(* IEC 61131-3 sources: rusty/tests/lit/single/functions, 19 files *)

(* ---- output_aggregate_initializers.st ---- *)
// RUN: %COMPILE %s && %RUN | %CHECK %s
// A struct literal, an array literal, and a string on a VAR_OUTPUT are applied by the lowered
// stack initializer of the function; the entry reset only zero-fills aggregates.
TYPE S : STRUCT
    x : INT;
    y : INT;
END_STRUCT END_TYPE

FUNCTION f
    VAR_OUTPUT
        out : S := (x := 7);
        arr : ARRAY[0..1] OF INT := [1, 2];
        s : STRING := 'abc';
    END_VAR
END_FUNCTION

FUNCTION main
    VAR
        v : S;
        a : ARRAY[0..1] OF INT;
        str : STRING;
    END_VAR
    v.y := 5;
    f(out => v, arr => a, s => str);
    printf('v = (%d, %d), a = [%d, %d], s = %s$N', v.x, v.y, a[0], a[1], str);
    // CHECK: v = (7, 0), a = [1, 2], s = abc
END_FUNCTION

(* ---- by_ref_argument_is_evaluated_once.st ---- *)
// RUN: %COMPILE %s && %RUN | %CHECK %s
// An expression passed to a by-reference input is evaluated once, also when the compiler carries it
// out through a replacement such as a builtin or a standard library call

VAR_GLOBAL
    calls : DINT;
END_VAR

FUNCTION next_number : DINT
    calls := calls + 1;
    next_number := calls;
END_FUNCTION

FUNCTION next_duration : TIME
    calls := calls + 1;
    next_duration := T#5s;
END_FUNCTION

FUNCTION read_number : DINT
VAR_INPUT {ref}
    in : DINT;
END_VAR
    read_number := in;
END_FUNCTION

FUNCTION read_duration : TIME
VAR_INPUT {ref}
    in : TIME;
END_VAR
    read_duration := in;
END_FUNCTION

FUNCTION main : DINT
    VAR
        n : DINT := 10;
        t : TIME := T#1s;
        result : DINT;
        duration : TIME;
    END_VAR

    result := read_number(n + next_number());
    printf('%d$N', result);                                                         // CHECK: 11
    printf('%d$N', calls);                                                          // CHECK: 1

    result := read_number(ADD(n, next_number()));
    printf('%d$N', result);                                                         // CHECK: 12
    printf('%d$N', calls);                                                          // CHECK: 2

    duration := read_duration(ADD(t, next_duration()));
    printf('%s$N', REF(TIME_TO_STRING(duration)));                                  // CHECK: T#6s
    printf('%d$N', calls);                                                          // CHECK: 3

END_FUNCTION

(* ---- call_with_array_access_on_result.st ---- *)
// RUN: %COMPILE %s && %RUN | %CHECK %s

FUNCTION foo: ARRAY[1..5] OF DINT
    foo := [5, 4, 3, 2, 1];
END_FUNCTION

FUNCTION alwaysOne: DINT
    alwaysOne := 1;
END_FUNCTION

FUNCTION main
    VAR
        value: DINT;
        one: DINT := 1;
        two: DINT := 2;
    END_VAR

    // CHECK: 5
    value := foo()[1];
    printf('%d$N', value);

    // CHECK: 3
    value := foo()[1 + 2];
    printf('%d$N', value);

    // CHECK: 5
    value := foo()[one];
    printf('%d$N', value);

    // CHECK: 3
    value := foo()[one + two];
    printf('%d$N', value);

    // CHECK: 5
    value := foo()[alwaysOne()];
    printf('%d$N', value);
END_FUNCTION

(* ---- deeply_nested_calls.st ---- *)
// RUN: %COMPILE %s && %RUN | %CHECK %s
// Deeply nested calls compile in time linear to their depth

FUNCTION increment : DINT
    VAR_INPUT
        value : DINT;
    END_VAR

    increment := value + 1;
END_FUNCTION

FUNCTION main
    VAR
        x : DINT := 0;
    END_VAR

    x := increment(increment(increment(increment(increment(increment(increment(increment(increment(increment(increment(increment(increment(increment(increment(increment(increment(increment(increment(increment(increment(increment(increment(increment(increment(increment(increment(increment(increment(increment(x))))))))))))))))))))))))))))));
    printf('%d$N', x);                                                              // CHECK: 30

END_FUNCTION

(* ---- default_params.st ---- *)
// RUN: %COMPILE %s && %RUN | %CHECK %s
FUNCTION func : int
  VAR_INPUT
    in : INT := 42;
  END_VAR
  func := in;
END_FUNCTION

FUNCTION main : DINT

    PRINTF('func complete:%d$N', func(13)); //CHECK: func complete:13
    PRINTF('func incomplete:%d$N', func()); //CHECK: func incomplete:42

END_FUNCTION

(* ---- function_output_should_be_cast_if_needed.st ---- *)
// RUN: %COMPILE %s && %RUN | %CHECK %s
FUNCTION outputCastIntToReal : INT
    VAR_OUTPUT
        result : REAL;
    END_VAR

    result := 42.0;
END_FUNCTION

FUNCTION outputNoCastInt : INT
    VAR_OUTPUT
        result : INT;
    END_VAR

    result := 52;
END_FUNCTION

FUNCTION outputCastRealToInt : INT
    VAR_OUTPUT
        result : INT;
    END_VAR

    result := 62;
END_FUNCTION

FUNCTION outputNoCastReal : INT
    VAR_OUTPUT
        result : REAL;
    END_VAR

    result := 72.0;
END_FUNCTION

FUNCTION main
    VAR
        i1 : INT;
        i2 : INT;
        r1 : REAL;
        r2 : REAL;
    END_VAR

    i1 := 31;
    i2 := 32;
    r1 := 33;
    r2 := 34;

    // ----------------- //
    // -- INT to REAL -- //

    outputCastIntToReal(
        result => i1
    );

    // CHECK: 42
    PRINTF('%d$N', i1);

    // ---------------- //
    // -- INT to INT -- //

    outputNoCastInt(
        result => i2
    );

    // CHECK: 52
    PRINTF('%d$N', i2);

    // ----------------- //
    // -- REAL to INT -- //

    outputCastRealToInt(
        result => r1
    );

    // CHECK: 62.0
    PRINTF('%.1f$N', r1);

    // ------------------ //
    // -- REAL to REAL -- //

    outputNoCastReal(
        result => r2
    );

    // CHECK: 72.0
    PRINTF('%.1f$N', r2);
END_FUNCTION

(* ---- function_parameter_with_bit_access.st ---- *)
// RUN: %COMPILE %s && %RUN | %CHECK %s
FUNCTION FLIP
    VAR_INPUT
        in: BYTE;
    END_VAR
    VAR_OUTPUT
        out : BYTE;
    END_VAR
    out := NOT(in);
END_FUNCTION

FUNCTION main
    VAR
        wordVar : WORD;
    END_VAR

    wordVar := 0;
    FLIP(2#01010101, wordVar.%b0);

    // CHECK: wordVar=170
    PRINTF('wordVar=%d$N', wordVar);
END_FUNCTION

(* ---- function_parameter_with_bit_access_named_params.st ---- *)
// RUN: %COMPILE %s && %RUN | %CHECK %s
FUNCTION FLIP
    VAR_INPUT
        in: BYTE;
    END_VAR
    VAR_OUTPUT
        out : BYTE;
    END_VAR
    out := NOT(in);
END_FUNCTION

FUNCTION main
    VAR
        wordVar : WORD;
    END_VAR

    wordVar := 0;
    FLIP(in := 2#01010101, out => wordVar.%b0);

    // CHECK: wordVar=170
    PRINTF('wordVar=%d$N', wordVar);
END_FUNCTION

(* ---- output_reset_on_every_call.st ---- *)
// RUN: %COMPILE %s && %RUN | %CHECK %s
// A function output that a path does not assign comes back at its default on every call, not at
// the value a previous call left in the caller's variable.
FUNCTION clamp_flag
    VAR_INPUT
        value : INT;
    END_VAR
    VAR_OUTPUT
        too_big : BOOL;
    END_VAR
    IF value > 2 THEN
        too_big := TRUE;
    END_IF
END_FUNCTION

FUNCTION main
    VAR
        i : INT;
        flag : BOOL;
    END_VAR
    FOR i := 1 TO 5 DO
        clamp_flag(i, flag);
        printf('%d: %d$N', i, flag);
    END_FOR
    // CHECK: 1: 0
    // CHECK-NEXT: 2: 0
    // CHECK-NEXT: 3: 1
    // CHECK-NEXT: 4: 1
    // CHECK-NEXT: 5: 1
    flag := TRUE;
    clamp_flag(1, flag);
    printf('after: %d$N', flag);
    // CHECK-NEXT: after: 0
END_FUNCTION

(* ---- function_block_output_should_be_cast_if_needed.st ---- *)
// RUN: %COMPILE %s && %RUN | %CHECK %s
FUNCTION_BLOCK outputCastIntToReal_fb
    VAR_OUTPUT
        result : REAL;
    END_VAR

    result := 42.0;
END_FUNCTION_BLOCK

FUNCTION_BLOCK outputNoCastInt_fb
    VAR_OUTPUT
        result : INT;
    END_VAR

    result := 52;
END_FUNCTION_BLOCK

FUNCTION_BLOCK outputCastRealToInt_fb
    VAR_OUTPUT
        result : INT;
    END_VAR

    result := 62;
END_FUNCTION_BLOCK

FUNCTION_BLOCK outputNoCastReal_fb
    VAR_OUTPUT
        result : REAL;
    END_VAR

    result := 72.0;
END_FUNCTION_BLOCK

FUNCTION main
    VAR
        outputCastIntToReal : outputCastIntToReal_fb;
        outputNoCastInt : outputNoCastInt_fb;
        outputCastRealToInt : outputCastRealToInt_fb;
        outputNoCastReal : outputNoCastReal_fb;

        i1 : INT;
        i2 : INT;
        r1 : REAL;
        r2 : REAL;
    END_VAR

    i1 := 31;
    i2 := 32;
    r1 := 33;
    r2 := 34;

    // ----------------- //
    // -- INT to REAL -- //

    outputCastIntToReal(
        result => i1
    );

    // CHECK: 42
    PRINTF('%d$N', i1);

    // ---------------- //
    // -- INT to INT -- //

    outputNoCastInt(
        result => i2
    );

    // CHECK: 52
    PRINTF('%d$N', i2);

    // ----------------- //
    // -- REAL to INT -- //

    outputCastRealToInt(
        result => r1
    );

    // CHECK: 62.0
    PRINTF('%.1f$N', r1);

    // ------------------ //
    // -- REAL to REAL -- //

    outputNoCastReal(
        result => r2
    );

    // CHECK: 72.0
    PRINTF('%.1f$N', r2);
END_FUNCTION

(* ---- function_output_to_bit_direct_access.st ---- *)
// RUN: %COMPILE %s && %RUN | %CHECK %s

// Regression test for https://github.com/PLC-lang/rusty/issues/1239
// `fun(out => bar.4)` and `myFb(out => bar.4)` previously generated IR that
// computed the bit address but never stored the function's output back into
// the underlying integer.
FUNCTION fun
    VAR_OUTPUT
        foo : BOOL;
    END_VAR
    foo := TRUE;
END_FUNCTION

FUNCTION_BLOCK fb
    VAR_OUTPUT
        foo : BOOL;
    END_VAR
    foo := TRUE;
END_FUNCTION_BLOCK

FUNCTION main : DINT
    VAR
        bar  : DINT;
        myFb : fb;
    END_VAR

    bar := 0;
    fun(foo => bar.4);
    PRINTF('after_fun=%d$N', bar);
    // CHECK: after_fun=16

    bar := 0;
    myFb(foo => bar.4);
    PRINTF('after_fb=%d$N', bar);
    // CHECK: after_fb=16

    // Non-zero seed: anchors that bits 0–3 are *preserved* when the FB output
    // writes bit 4. A regression that clobbered the integer (e.g. wrote a full
    // word instead of just the bit) would surface here as 16 instead of 17.
    bar := 1;
    myFb(foo => bar.4);
    PRINTF('after_fb_seeded=%d$N', bar);
    // CHECK: after_fb_seeded=17
END_FUNCTION

(* ---- output_pointer_type_default.st ---- *)
// RUN: %COMPILE %s && %RUN | %CHECK %s
// A pointer-typed output keeps its constructor call, so an address-valued default of its type,
// which codegen cannot store as a constant, is applied on every call.
VAR_GLOBAL
    g : DINT := 99;
END_VAR

TYPE P : POINTER TO DINT := ADR(g); END_TYPE

FUNCTION_BLOCK Fb
    METHOD m
        VAR_OUTPUT
            out : P;
        END_VAR
    END_METHOD
END_FUNCTION_BLOCK

FUNCTION f
    VAR_OUTPUT
        out : P;
    END_VAR
END_FUNCTION

FUNCTION main
    VAR
        fb : Fb;
        p : P;
    END_VAR
    p := ADR(p);
    f(out => p);
    printf('function: out^ = %d, out = ADR(g): %d$N', p^, p = ADR(g));
    // CHECK: function: out^ = 99, out = ADR(g): 1

    p := ADR(p);
    fb.m(out => p);
    printf('method: out^ = %d, out = ADR(g): %d$N', p^, p = ADR(g));
    // CHECK-NEXT: method: out^ = 99, out = ADR(g): 1
END_FUNCTION

(* ---- output_scalar_address_default.st ---- *)
// RUN: %COMPILE %s && %RUN | %CHECK %s
// A scalar type whose default is an address, which codegen cannot store as a constant, is applied
// to an output of that type by the type's constructor on every call, in a function and a method.
VAR_GLOBAL
    g : DINT := 99;
END_VAR

TYPE A : LWORD := ADR(g); END_TYPE

FUNCTION_BLOCK Fb
    METHOD m
        VAR_OUTPUT
            out : A;
        END_VAR
    END_METHOD
END_FUNCTION_BLOCK

FUNCTION f
    VAR_OUTPUT
        out : A;
    END_VAR
END_FUNCTION

FUNCTION main
    VAR
        fb : Fb;
        a : A;
    END_VAR
    a := 1;
    f(out => a);
    printf('function: out = ADR(g): %d$N', a = ADR(g));
    // CHECK: function: out = ADR(g): 1

    a := 1;
    fb.m(out => a);
    printf('method: out = ADR(g): %d$N', a = ADR(g));
    // CHECK-NEXT: method: out = ADR(g): 1
END_FUNCTION

(* ---- output_scalar_type_defaults.st ---- *)
// RUN: %COMPILE %s && %RUN | %CHECK %s
// Outputs of an alias, subrange, enum, or struct type start every call at the default of their
// type, in a function and in a method alike. A scalar output needs no constructor call, so an
// alias of an elementary type must compile as an output.
TYPE MyInt : INT; END_TYPE
TYPE Preset : DINT := 20; END_TYPE
TYPE Pct : INT(0..100) := 50; END_TYPE
TYPE Color : (Red, Green := 5, Blue) := Green; END_TYPE
TYPE S : STRUCT
    a : INT := 7;
END_STRUCT END_TYPE

FUNCTION_BLOCK Fb
    METHOD m
        VAR_OUTPUT
            p : MyInt;
            q : Preset;
            r : Pct;
            c : Color;
            st : S;
        END_VAR
    END_METHOD
END_FUNCTION_BLOCK

FUNCTION f
    VAR_OUTPUT
        p : MyInt;
        q : Preset;
        r : Pct;
        c : Color;
        st : S;
    END_VAR
END_FUNCTION

FUNCTION main
    VAR
        fb : Fb;
        a : MyInt;
        b : Preset;
        r : Pct;
        c : Color;
        st : S;
    END_VAR
    a := 1; b := 1; r := 1; c := Blue; st.a := 1;
    f(p => a, q => b, r => r, c => c, st => st);
    printf('function: a = %d, b = %d, r = %d, c = %d, st.a = %d$N', a, b, r, c, st.a);
    // CHECK: function: a = 0, b = 20, r = 50, c = 5, st.a = 7

    a := 1; b := 1; r := 1; c := Blue; st.a := 1;
    fb.m(p => a, q => b, r => r, c => c, st => st);
    printf('method: a = %d, b = %d, r = %d, c = %d, st.a = %d$N', a, b, r, c, st.a);
    // CHECK-NEXT: method: a = 0, b = 20, r = 50, c = 5, st.a = 7
END_FUNCTION

(* ---- segmented_variable_blocks_with_implicit_arguments_call.st ---- *)
// RUN: %COMPILE %s && %RUN | %CHECK %s

FUNCTION_BLOCK foo
    VAR
        placeholder_one: DINT;
    END_VAR

    VAR_INPUT
        a, b: DINT;
    END_VAR

    VAR
        placeholder_two: DINT;
    END_VAR

    VAR_OUTPUT
        c: DINT;
    END_VAR

    c := a + b;
END_FUNCTION_BLOCK

FUNCTION main
    VAR
        foo: foo;
        local_a, local_b, local_c: DINT := 2;
    END_VAR

    foo(local_a, local_b, local_c);
    printf('%d$N', local_c); // CHECK: 4
END_FUNCTION

(* ---- function_output_declared_as_plain_string_with_aggregate_return_type_should_evaluate_correctly.st ---- *)
// RUN: %COMPILE %s && %RUN | %CHECK %s
FUNCTION F : STRING
    VAR_INPUT
        Key : STRING[1023];
    END_VAR
    VAR_OUTPUT
        Value : STRING;
    END_VAR

    Value := 'AAAAAAAAAAAAAAAAAAAAAAAAAAAAAAAAAAAAAAAAAAAAAAAAAAAAAAAAAAAAAAAAAAAAAAAAAAAAAAAAAAAAAAAAAAAAAAAAAAAAAAAAAAAAAAAAAAAAAAAAAAAAAAAAAAAAAAAAAAAAAAAAAAAAAAAAAAAAAAAAAAAAAAAAAAAAAAAAAAAAAAAAAAAAAAAAAAAAAAAAAAAAAAAAAAAAAAAAAAAAAAAAAAAAAAAAAAAAAAAAAAAAAAAAAAAAAAAAAAAAAAAAAAAAAAAAAAAAAAAAAAAAAAAAAAAAAAAAAAAAAAAAAAAAAAAAAAAAAAAAAAAAAAAAAAAAAAAAAAAAAAAAAAAAAAAAAAAAAAAAAAAAAAAAAAAAAAAAAAAAAAAAAAAAAAAAAAAAAAAAAAAAAAAAAAAAAAAAAAAAAAAAAAAAAAAAAAAAAAAAAAAAAAAAAAAAAAAAAAAAAAAAAAAAAAAAAAAAAAAAAAAAAAAAAAAAAAAAAAAAAAAAAAAAAAAAAAAAAAAAAAAAAAAAAAAAAAAAAAAAAAAAAAAAAAAAAAAAAAAAAAAAAAAAAAAAAAAAAAAAAAAAAAAAAAAAAAAAAAAAAAAAAAAAAAAAAAAAAAAAAAAAAAAAAAAAAAAAAAAAAAAAAAAAAAAAAAAAAAAAAAAAAAAAAAAAAAAAAAAAAAAAAAAAAAAAAAAAAAAAAAAAAAAAAAAAAAAAAAAAAAAAAAAAAAAAAAAAAAAAAAAAAAAAAAAAAAAAAAAAAAAAAAAAAAAAAAAAAAAAAAAAAAAAAAAAAAAAAAAAAAAAAAAAAAAAAAAAAAAAAAAAAAAAAAAAAAAAAAAAAAAAAAAAAAAAAAAAAAAAAAAAAAAAAAAAAAAAAAAAAAAAAAAAAAAAAAAAAAAAAAAAAAAAAAAAAAAAAAAAAAAAAAAAAAAAAAAAAAAAAAAAAAAAAAAAAAAAAAAAAAAAAAAAAAAAAAAAAAAAAAAAAAAAAAAAAAAAAAAAAAAAAAAAAAAAAAAAAAAAAAA';
    F := 'returned';
END_FUNCTION

PROGRAM mainProg
    VAR
        MyString : STRING;          // too-small caller buffer
        MyInt    : INT  := 1234;    // guards
        MyGuard  : DINT := 24681357;
        retString : STRING;
    END_VAR
    retString := F('key', MyString);

    // CHECK: ret=returned my_int=1234 my_guard=24681357 value_prefix=AAAAAAAA
    printf('ret=%.8s my_int=%d my_guard=%d value_prefix=%.8s$N', retString, MyInt, MyGuard, MyString);
END_PROGRAM

FUNCTION main : DINT
    mainProg();
END_FUNCTION

(* ---- function_output_should_be_ignored_if_unassigned.st ---- *)
// RUN: %COMPILE %s && %RUN | %CHECK %s
FUNCTION GetVal : DINT
    VAR_OUTPUT
        Value : STRING[80];
    END_VAR

    Value := 'Hello World';

    GetVal := 2;
END_FUNCTION

PROGRAM mainProg
    VAR
        s : STRING;
    END_VAR

    // CHECK: 2
    IF GetVal(Value => ) = 0 THEN
        PRINTF('0$N');
    ELSE
        PRINTF('2$N');
    END_IF
END_PROGRAM

FUNCTION main
    mainProg();
END_FUNCTION

(* ---- function_output_should_truncate_when_string_sizes_are_mismatched.st ---- *)
// RUN: %COMPILE %s && %RUN | %CHECK %s
FUNCTION Config_GetString : DINT
    VAR_INPUT
        Key : STRING[1023];
    END_VAR
    VAR_OUTPUT
        Value : STRING[28];
    END_VAR

    Value := 'I am a non-truncated string';

END_FUNCTION

FUNCTION Config_GetString_Auto : DINT
    VAR_INPUT
        Key : STRING[1023];
    END_VAR
    VAR_OUTPUT
        Value : STRING;
    END_VAR

    Value := 'I am an automatically sized non-truncated string';

END_FUNCTION

PROGRAM mainProg
    VAR
        MyString : STRING[10];
        MyInt: INT := 1234;
        retValue : DINT;
    END_VAR

    retValue := Config_GetString('/some/config/value', MyString);

    // CHECK: I am a non
    PRINTF('%s$N', MyString);

    retValue := Config_GetString_Auto('/some/config/value', MyString);

    // CHECK: I am an au
    PRINTF('%s$N', MyString);
END_PROGRAM

FUNCTION main
    mainProg();
END_FUNCTION

(* ---- function_output_with_aggregate_return_type_should_evaluate_correctly.st ---- *)
// RUN: %COMPILE %s && %RUN | %CHECK %s
FUNCTION F : STRING
    VAR_INPUT
        Key : STRING[1023];
    END_VAR
    VAR_OUTPUT
        Value : STRING[1023];
    END_VAR

    Value := 'AAAAAAAAAAAAAAAAAAAAAAAAAAAAAAAAAAAAAAAAAAAAAAAAAAAAAAAAAAAAAAAAAAAAAAAAAAAAAAAAAAAAAAAAAAAAAAAAAAAAAAAAAAAAAAAAAAAAAAAAAAAAAAAAAAAAAAAAAAAAAAAAAAAAAAAAAAAAAAAAAAAAAAAAAAAAAAAAAAAAAAAAAAAAAAAAAAAAAAAAAAAAAAAAAAAAAAAAAAAAAAAAAAAAAAAAAAAAAAAAAAAAAAAAAAAAAAAAAAAAAAAAAAAAAAAAAAAAAAAAAAAAAAAAAAAAAAAAAAAAAAAAAAAAAAAAAAAAAAAAAAAAAAAAAAAAAAAAAAAAAAAAAAAAAAAAAAAAAAAAAAAAAAAAAAAAAAAAAAAAAAAAAAAAAAAAAAAAAAAAAAAAAAAAAAAAAAAAAAAAAAAAAAAAAAAAAAAAAAAAAAAAAAAAAAAAAAAAAAAAAAAAAAAAAAAAAAAAAAAAAAAAAAAAAAAAAAAAAAAAAAAAAAAAAAAAAAAAAAAAAAAAAAAAAAAAAAAAAAAAAAAAAAAAAAAAAAAAAAAAAAAAAAAAAAAAAAAAAAAAAAAAAAAAAAAAAAAAAAAAAAAAAAAAAAAAAAAAAAAAAAAAAAAAAAAAAAAAAAAAAAAAAAAAAAAAAAAAAAAAAAAAAAAAAAAAAAAAAAAAAAAAAAAAAAAAAAAAAAAAAAAAAAAAAAAAAAAAAAAAAAAAAAAAAAAAAAAAAAAAAAAAAAAAAAAAAAAAAAAAAAAAAAAAAAAAAAAAAAAAAAAAAAAAAAAAAAAAAAAAAAAAAAAAAAAAAAAAAAAAAAAAAAAAAAAAAAAAAAAAAAAAAAAAAAAAAAAAAAAAAAAAAAAAAAAAAAAAAAAAAAAAAAAAAAAAAAAAAAAAAAAAAAAAAAAAAAAAAAAAAAAAAAAAAAAAAAAAAAAAAAAAAAAAAAAAAAAAAAAAAAAAAAAAAAAAAAAAAAAAAAAAAAAAAAAAAAAAAAAAAAAAAAAAAAAAAAAAAAAAAAA';
    F := 'returned';
END_FUNCTION

PROGRAM mainProg
    VAR
        MyString : STRING;          // too-small caller buffer
        MyInt    : INT  := 1234;    // guards
        MyGuard  : DINT := 24681357;
        retString : STRING;
    END_VAR
    retString := F('key', MyString);

    // CHECK: ret=returned my_int=1234 my_guard=24681357 value_prefix=AAAAAAAA
    printf('ret=%.8s my_int=%d my_guard=%d value_prefix=%.8s$N', retString, MyInt, MyGuard, MyString);
END_PROGRAM

FUNCTION main : DINT
    mainProg();
END_FUNCTION
